// TIA Portal V21 export
// export: Created 2026-08-21T20:18:51.5900179Z, ExportSetting None, DisplayName Totally Integrated Automation Portal, DisplayVersion V21, DisplayName STEP 7 Professional, DisplayVersion V21, DisplayName STEP 7 Safety, DisplayVersion V21, DisplayName Tech WebApplication, DisplayVersion V21, DisplayName WinCC Basic/Comfort/Advanced, DisplayVersion V21, DisplayName WinCC Professional, DisplayVersion V21, DisplayName WinCC Unified, DisplayVersion V21
DATA_BLOCK "P100_Type"   // DB3
// stored: InstanceOfName MTPMonBinDrv_Type1, InstanceOfType FB
"MTPMonBinDrv_Type1"
   // VAR_INPUT
   //    from_Ctrl { ExternalAccessible := 'False'; ExternalVisible := 'False'; ExternalWritable := 'False'} : "StruCm";
   //    Service_Occupied { ExternalAccessible := 'False'; ExternalVisible := 'False'; ExternalWritable := 'False'} : Bool;
   //    Cmd_Auto { ExternalAccessible := 'False'; ExternalVisible := 'False'; ExternalWritable := 'False'} : Bool;
   //    Cmd_Man { ExternalAccessible := 'False'; ExternalVisible := 'False'; ExternalWritable := 'False'} : Bool;
   //    Cmd_StartAut { ExternalAccessible := 'False'; ExternalVisible := 'False'; ExternalWritable := 'False'} : Bool;
   //    Cmd_StopAut { ExternalAccessible := 'False'; ExternalVisible := 'False'; ExternalWritable := 'False'} : Bool;
   //    Cmd_Reset { ExternalAccessible := 'False'; ExternalVisible := 'False'; ExternalWritable := 'False'} : Bool;
   //    PV_In : Bool;
   //    Intlk04_In01 { ExternalAccessible := 'False'; ExternalVisible := 'False'; ExternalWritable := 'False'} : "DigVal";
   //    Intlk04_InvIn01 : Bool;
   //    Intlk04_In1String : String;
   //    Intlk04_In02 { ExternalAccessible := 'False'; ExternalVisible := 'False'; ExternalWritable := 'False'} : "DigVal";
   //    Intlk04_InvIn02 : Bool;
   //    Intlk04_In2String { ExternalAccessible := 'False'; ExternalVisible := 'False'; ExternalWritable := 'False'} : String;
   //    Intlk04_In03 { ExternalAccessible := 'False'; ExternalVisible := 'False'; ExternalWritable := 'False'} : "DigVal";
   //    Intlk04_InvIn03 : Bool;
   //    Intlk04_In3String { ExternalAccessible := 'False'; ExternalVisible := 'False'; ExternalWritable := 'False'} : String;
   //    Intlk04_In04 { ExternalAccessible := 'False'; ExternalVisible := 'False'; ExternalWritable := 'False'} : "DigVal";
   //    Intlk04_InvIn04 : Bool;
   //    Intlk04_In4String { ExternalAccessible := 'False'; ExternalVisible := 'False'; ExternalWritable := 'False'} : String;
   // END_VAR
   // VAR_OUTPUT
   //    to_Ctrl { ExternalAccessible := 'False'; ExternalVisible := 'False'; ExternalWritable := 'False'} : "StruCm";
   //    Occupied { ExternalAccessible := 'False'; ExternalVisible := 'False'; ExternalWritable := 'False'} : Bool;
   //    AutAct { ExternalAccessible := 'False'; ExternalVisible := 'False'; ExternalWritable := 'False'} : Bool;
   //    ManAct { ExternalAccessible := 'False'; ExternalVisible := 'False'; ExternalWritable := 'False'} : Bool;
   //    PV_Out { ExternalAccessible := 'False'; ExternalVisible := 'False'; ExternalWritable := 'False'} : Bool;
   //    FbkRunOut : Bool;
   //    RunOut : Bool;
   //    Stop { ExternalAccessible := 'False'; ExternalVisible := 'False'; ExternalWritable := 'False'} : Bool;
   //    GrpErr { ExternalAccessible := 'False'; ExternalVisible := 'False'; ExternalWritable := 'False'} : Bool;
   // END_VAR
   // VAR
   //    ChOut { S7_SetPoint := 'True'} : "DiOu";
   //    DiChIn { S7_SetPoint := 'True'} : "DiIn";
   //    Intlk04_IDB : "Intlk04";
   //    MotL_IDB { S7_SetPoint := 'True'} : "MotL";
   //    MTPMonBinDrv_IDB { ExternalVisible := 'False'; S7_SetPoint := 'True'} : "MTPMonBinDrv";
   // END_VAR
BEGIN
   Intlk04_IDB.DataHMI.In01_Text := '';
   Intlk04_IDB.DataHMI.BypIn01 := FALSE;
   Intlk04_IDB.DataHMI.AV01 := 0.0;
   Intlk04_IDB.DataHMI.AV01_Unit := 0;
   Intlk04_IDB.DataHMI.In02_Text := '';
   Intlk04_IDB.DataHMI.BypIn02 := FALSE;
   Intlk04_IDB.DataHMI.AV02 := 0.0;
   Intlk04_IDB.DataHMI.AV02_Unit := 0;
   Intlk04_IDB.DataHMI.In03_Text := '';
   Intlk04_IDB.DataHMI.BypIn03 := FALSE;
   Intlk04_IDB.DataHMI.AV03 := 0.0;
   Intlk04_IDB.DataHMI.AV03_Unit := 0;
   Intlk04_IDB.DataHMI.In04_Text := '';
   Intlk04_IDB.DataHMI.BypIn04 := FALSE;
   Intlk04_IDB.DataHMI.AV04 := 0.0;
   Intlk04_IDB.DataHMI.AV04_Unit := 0;
   Intlk04_IDB.DataHMI.RstOp := FALSE;
   Intlk04_IDB.DataHMI.RstBypOp := FALSE;
   Intlk04_IDB.DataHMI.OS_PermOut := 16#FFFF_FFFF;
   Intlk04_IDB.DataHMI.OS_PermLog := 16#FFF0_FFF9;
   Intlk04_IDB.DataHMI.OpSt_Out := 16#0000_0000;
   Intlk04_IDB.DataHMI.ST_Worst := 16#80;
   Intlk04_IDB.DataHMI.Status1 := 16#0000_0202;
   Intlk04_IDB.DataHMI.Status2 := 16#0000_000E;
   Intlk04_IDB.DataHMI.Status3 := 16#0000_0000;
   Intlk04_IDB.DataHMI.Status4 := 16#0000_000E;
   Intlk04_IDB.DataHMI.Status5 := 16#0000_0000;
   Intlk04_IDB.DataHMI.Status6 := 16#0000_0000;
   Intlk04_IDB.DataHMI.Status7 := 16#0000_000F;
   Intlk04_IDB.DataHMI.Status8 := 16#0000_0000;
   MotL_IDB.Monitor := TRUE;
   MotL_IDB.MonTiStatic := 10.0;
   MotL_IDB.MonTiDynamic := 10.0;
   MotL_IDB.MonTiDyStop := 3.0;
   MotL_IDB.SimOn := FALSE;
   MotL_IDB.DataHMI.StartMan := FALSE;
   MotL_IDB.DataHMI.StopMan := FALSE;
   MotL_IDB.DataHMI.AutModOp := FALSE;
   MotL_IDB.DataHMI.ManModOp := FALSE;
   MotL_IDB.DataHMI.LocalOp := FALSE;
   MotL_IDB.DataHMI.OosOp := FALSE;
   MotL_IDB.DataHMI.LocalLi := FALSE;
   MotL_IDB.DataHMI.StartLocal := FALSE;
   MotL_IDB.DataHMI.StopLocal := FALSE;
   MotL_IDB.DataHMI.Monitor := TRUE;
   MotL_IDB.DataHMI.MonTiStatic := 10.0;
   MotL_IDB.DataHMI.MonTiDynamic := 10.0;
   MotL_IDB.DataHMI.MonTiDyStop := 3.0;
   MotL_IDB.DataHMI.RapidStp := FALSE;
   MotL_IDB.DataHMI.RstOp := FALSE;
   MotL_IDB.DataHMI.Permit_ST := 16#FF;
   MotL_IDB.DataHMI.Intlock_ST := 16#80;
   MotL_IDB.DataHMI.Protect_ST := 16#FF;
   MotL_IDB.DataHMI.CurrMon := 0;
   MotL_IDB.DataHMI.FbkRunOut := FALSE;
   MotL_IDB.DataHMI.OS_PermOut := 16#FFFF_FFFF;
   MotL_IDB.DataHMI.OS_PermLog := 16#7BFF_FF49;
   MotL_IDB.DataHMI.OpSt_Out := 16#0000_0000;
   MotL_IDB.DataHMI.ST_Worst := 16#80;
   MotL_IDB.DataHMI.Status1 := 16#1081_0280;
   MotL_IDB.DataHMI.Status2 := 16#4010_0000;
   MotL_IDB.DataHMI.Status3 := 16#0200_8000;
   MotL_IDB.DataHMI.Status4 := 16#0000_0400;
   MotL_IDB.DataHMI.AlarmState := 16#0000;
   MotL_IDB.Start.Value := FALSE;
   MotL_IDB.Start.InternalUseBit1 := FALSE;
   MotL_IDB.Start.InternalUseBit2 := FALSE;
   MotL_IDB.Start.InternalUseBit3 := FALSE;
   MotL_IDB.Start.InternalUseBit4 := FALSE;
   MotL_IDB.Start.InternalUseBit5 := FALSE;
   MotL_IDB.Start.InternalUseBit6 := FALSE;
   MotL_IDB.Start.InternalUseBit7 := FALSE;
   MotL_IDB.Start.ST := 16#80;
   MotL_IDB.LocalAct.Value := FALSE;
   MotL_IDB.LocalAct.InternalUseBit1 := FALSE;
   MotL_IDB.LocalAct.InternalUseBit2 := FALSE;
   MotL_IDB.LocalAct.InternalUseBit3 := FALSE;
   MotL_IDB.LocalAct.InternalUseBit4 := FALSE;
   MotL_IDB.LocalAct.InternalUseBit5 := FALSE;
   MotL_IDB.LocalAct.InternalUseBit6 := FALSE;
   MotL_IDB.LocalAct.InternalUseBit7 := FALSE;
   MotL_IDB.LocalAct.ST := 16#80;
   MotL_IDB.AutAct.Value := FALSE;
   MotL_IDB.AutAct.InternalUseBit1 := FALSE;
   MotL_IDB.AutAct.InternalUseBit2 := FALSE;
   MotL_IDB.AutAct.InternalUseBit3 := FALSE;
   MotL_IDB.AutAct.InternalUseBit4 := FALSE;
   MotL_IDB.AutAct.InternalUseBit5 := FALSE;
   MotL_IDB.AutAct.InternalUseBit6 := FALSE;
   MotL_IDB.AutAct.InternalUseBit7 := FALSE;
   MotL_IDB.AutAct.ST := 16#80;
   MotL_IDB.ManAct.Value := TRUE;
   MotL_IDB.ManAct.InternalUseBit1 := FALSE;
   MotL_IDB.ManAct.InternalUseBit2 := FALSE;
   MotL_IDB.ManAct.InternalUseBit3 := FALSE;
   MotL_IDB.ManAct.InternalUseBit4 := FALSE;
   MotL_IDB.ManAct.InternalUseBit5 := FALSE;
   MotL_IDB.ManAct.InternalUseBit6 := FALSE;
   MotL_IDB.ManAct.InternalUseBit7 := FALSE;
   MotL_IDB.ManAct.ST := 16#80;
   MotL_IDB.OosAct.Value := FALSE;
   MotL_IDB.OosAct.InternalUseBit1 := FALSE;
   MotL_IDB.OosAct.InternalUseBit2 := FALSE;
   MotL_IDB.OosAct.InternalUseBit3 := FALSE;
   MotL_IDB.OosAct.InternalUseBit4 := FALSE;
   MotL_IDB.OosAct.InternalUseBit5 := FALSE;
   MotL_IDB.OosAct.InternalUseBit6 := FALSE;
   MotL_IDB.OosAct.InternalUseBit7 := FALSE;
   MotL_IDB.OosAct.ST := 16#80;
   MotL_IDB.Run.Value := FALSE;
   MotL_IDB.Run.InternalUseBit1 := FALSE;
   MotL_IDB.Run.InternalUseBit2 := FALSE;
   MotL_IDB.Run.InternalUseBit3 := FALSE;
   MotL_IDB.Run.InternalUseBit4 := FALSE;
   MotL_IDB.Run.InternalUseBit5 := FALSE;
   MotL_IDB.Run.InternalUseBit6 := FALSE;
   MotL_IDB.Run.InternalUseBit7 := FALSE;
   MotL_IDB.Run.ST := 16#80;
   MotL_IDB.Stop.Value := TRUE;
   MotL_IDB.Stop.InternalUseBit1 := FALSE;
   MotL_IDB.Stop.InternalUseBit2 := FALSE;
   MotL_IDB.Stop.InternalUseBit3 := FALSE;
   MotL_IDB.Stop.InternalUseBit4 := FALSE;
   MotL_IDB.Stop.InternalUseBit5 := FALSE;
   MotL_IDB.Stop.InternalUseBit6 := FALSE;
   MotL_IDB.Stop.InternalUseBit7 := FALSE;
   MotL_IDB.Stop.ST := 16#80;
   MotL_IDB.SrMonTime := 10.0;
   MotL_IDB.SxFirstStart := FALSE;
   MotL_IDB.SxCmdStart := FALSE;
   MotL_IDB.SxLastMode := FALSE;
END_DATA_BLOCK
